// TIA Portal V19 export
FUNCTION_BLOCK "V20_BLOCK"   // FB40, LAD
{ S7_Optimized_Access := 'FALSE' }
// stored: SetENOAutomatically false
   VAR
      MB_LOAD { S7_SetPoint := 'True'} : Modbus_Comm_Load;
      MB_READ_ZSW { S7_SetPoint := 'True'} : Modbus_Master;
      MB_READ_HIW { S7_SetPoint := 'True'} : Modbus_Master;
      MB_WRITE_STW { S7_SetPoint := 'True'} : Modbus_Master;
      MB_WRITE_HSW { S7_SetPoint := 'True'} : Modbus_Master;
      DRIVE { S7_SetPoint := 'True'} : Array[1..11] of "VFD";
      DRIVE_ID { S7_SetPoint := 'True'} : Int := 1;
      STATUS : Int;
      MB_DB : P2P_MB_BASE;
      ZSW_DELAY { S7_SetPoint := 'True'} : TON_TIME;
      HIW_DELAY { S7_SetPoint := 'True'} : TON_TIME;
      STW_DELAY { S7_SetPoint := 'True'} : TON_TIME;
      HSW_DELAY { S7_SetPoint := 'True'} : TON_TIME;
      MB_READ_DI { S7_SetPoint := 'True'} : Modbus_Master;
      Modbus_Master_Instance { S7_SetPoint := 'True'} : Modbus_Master;
   END_VAR
   // DRIVE[1].ADDR := 1;
   // DRIVE[2].ADDR := 2;
   // DRIVE[3].ADDR := 3;
   // DRIVE[4].ADDR := 4;
   // DRIVE[5].ADDR := 5;
   // DRIVE[6].ADDR := 6;
   VAR_TEMP   // added for the SCL form of the ladder/FBD networks
      _w1 : Bool;
   END_VAR
BEGIN

REGION Network 1
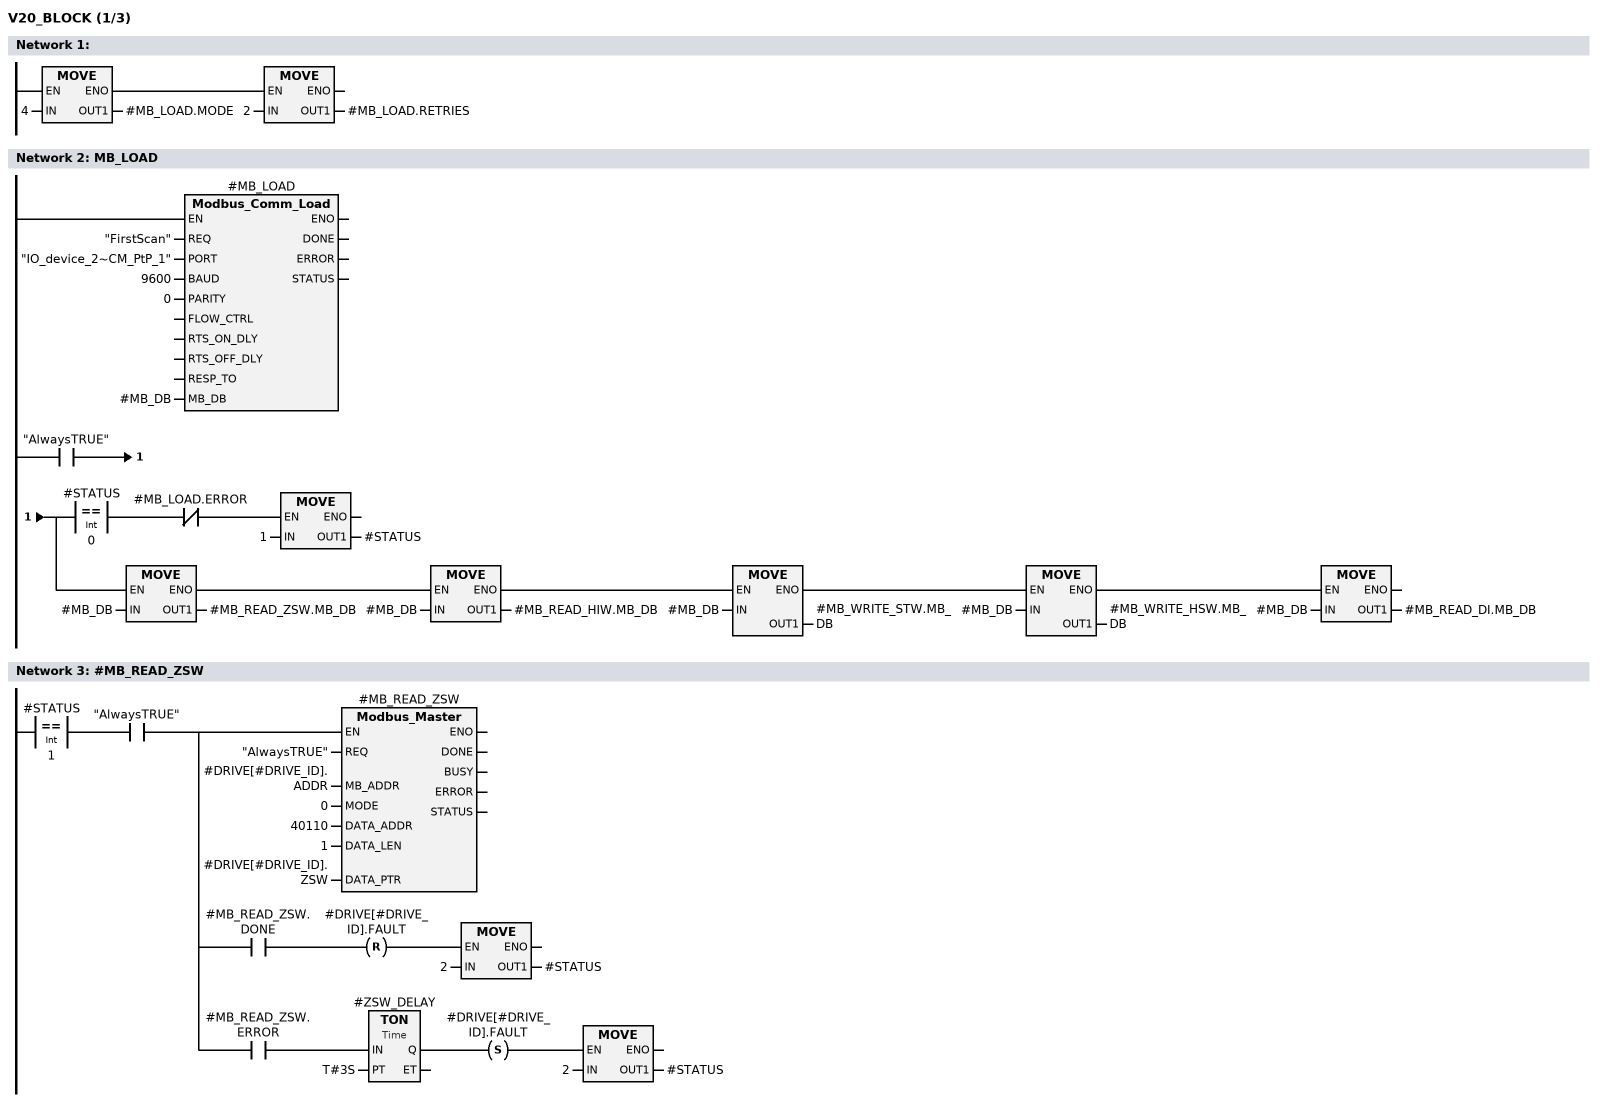
   RUNG wire#powerrail
      Move(in := 4, out1 => #MB_LOAD.MODE)
      Move(in := 2, out1 => #MB_LOAD.RETRIES)
   END_RUNG
   // the same network as SCL:
   #MB_LOAD.MODE := 4;
   #MB_LOAD.RETRIES := 2;
END_REGION

REGION Network 2: MB_LOAD
   RUNG wire#powerrail
      #MB_LOAD.Modbus_Comm_Load(REQ := "FirstScan", PORT := "IO_device_2~CM_PtP_1", BAUD := 9600, PARITY := 0, FLOW_CTRL :=, RTS_ON_DLY :=, RTS_OFF_DLY :=, RESP_TO :=, MB_DB := #MB_DB, DONE =>, ERROR =>, STATUS =>)
   END_RUNG
   RUNG wire#powerrail
      Contact( "AlwaysTRUE" )
      wire#w1
      { S7_Templates := "SrcType := Int" } EQ_Contact(in1 := #STATUS, in2 := 0)
      I_Contact( #MB_LOAD.ERROR )
      Move(in := 1, out1 => #STATUS)
   END_RUNG
   RUNG wire#w1
      Move(in := #MB_DB, out1 => #MB_READ_ZSW.MB_DB)
      Move(in := #MB_DB, out1 => #MB_READ_HIW.MB_DB)
      Move(in := #MB_DB, out1 => #MB_WRITE_STW.MB_DB)
      Move(in := #MB_DB, out1 => #MB_WRITE_HSW.MB_DB)
      Move(in := #MB_DB, out1 => #MB_READ_DI.MB_DB)
   END_RUNG
   // the same network as SCL:
   #MB_LOAD(REQ := "FirstScan", PORT := "IO_device_2~CM_PtP_1", BAUD := 9600, PARITY := 0, MB_DB := #MB_DB);   // Modbus_Comm_Load
   IF "AlwaysTRUE" AND (#STATUS = 0) AND NOT #MB_LOAD.ERROR THEN #STATUS := 1; END_IF;
   IF "AlwaysTRUE" THEN
       #MB_READ_ZSW.MB_DB := #MB_DB;
       #MB_READ_HIW.MB_DB := #MB_DB;
       #MB_WRITE_STW.MB_DB := #MB_DB;
       #MB_WRITE_HSW.MB_DB := #MB_DB;
       #MB_READ_DI.MB_DB := #MB_DB;
   END_IF;
END_REGION

REGION Network 3: #MB_READ_ZSW
   RUNG wire#powerrail
      { S7_Templates := "SrcType := Int" } EQ_Contact(in1 := #STATUS, in2 := 1)
      Contact( "AlwaysTRUE" )
      wire#w1
      #MB_READ_ZSW.Modbus_Master(REQ := "AlwaysTRUE", MB_ADDR := #DRIVE[#DRIVE_ID].ADDR, MODE := 0, DATA_ADDR := 40110, DATA_LEN := 1, DATA_PTR := #DRIVE[#DRIVE_ID].ZSW, DONE =>, BUSY =>, ERROR =>, STATUS =>)
   END_RUNG
   RUNG wire#w1
      Contact( #MB_READ_ZSW.DONE )
      R_Coil( #DRIVE[#DRIVE_ID].FAULT )
      Move(in := 2, out1 => #STATUS)
   END_RUNG
   RUNG wire#w1
      Contact( #MB_READ_ZSW.ERROR )
      { S7_Templates := "time_type := Time" } #ZSW_DELAY.TON(pt := T#3S, et =>)
      S_Coil( #DRIVE[#DRIVE_ID].FAULT )
      Move(in := 2, out1 => #STATUS)
   END_RUNG
   // the same network as SCL:
   #_w1 := (#STATUS = 1) AND "AlwaysTRUE";
   IF #_w1 THEN
       #MB_READ_ZSW(REQ := "AlwaysTRUE",   // Modbus_Master
                    MB_ADDR := #DRIVE[#DRIVE_ID].ADDR,
                    MODE := 0,
                    DATA_ADDR := 40110,
                    DATA_LEN := 1,
                    DATA_PTR := #DRIVE[#DRIVE_ID].ZSW);
   END_IF;
   IF #_w1 AND #MB_READ_ZSW.DONE THEN
       #DRIVE[#DRIVE_ID].FAULT := FALSE;
       #STATUS := 2;
   END_IF;
   #ZSW_DELAY(IN := #_w1 AND #MB_READ_ZSW.ERROR, PT := T#3S);   // TON
   IF #ZSW_DELAY.Q THEN
       #DRIVE[#DRIVE_ID].FAULT := TRUE;
       #STATUS := 2;
   END_IF;
END_REGION

REGION Network 4: #MB_READ_HIW
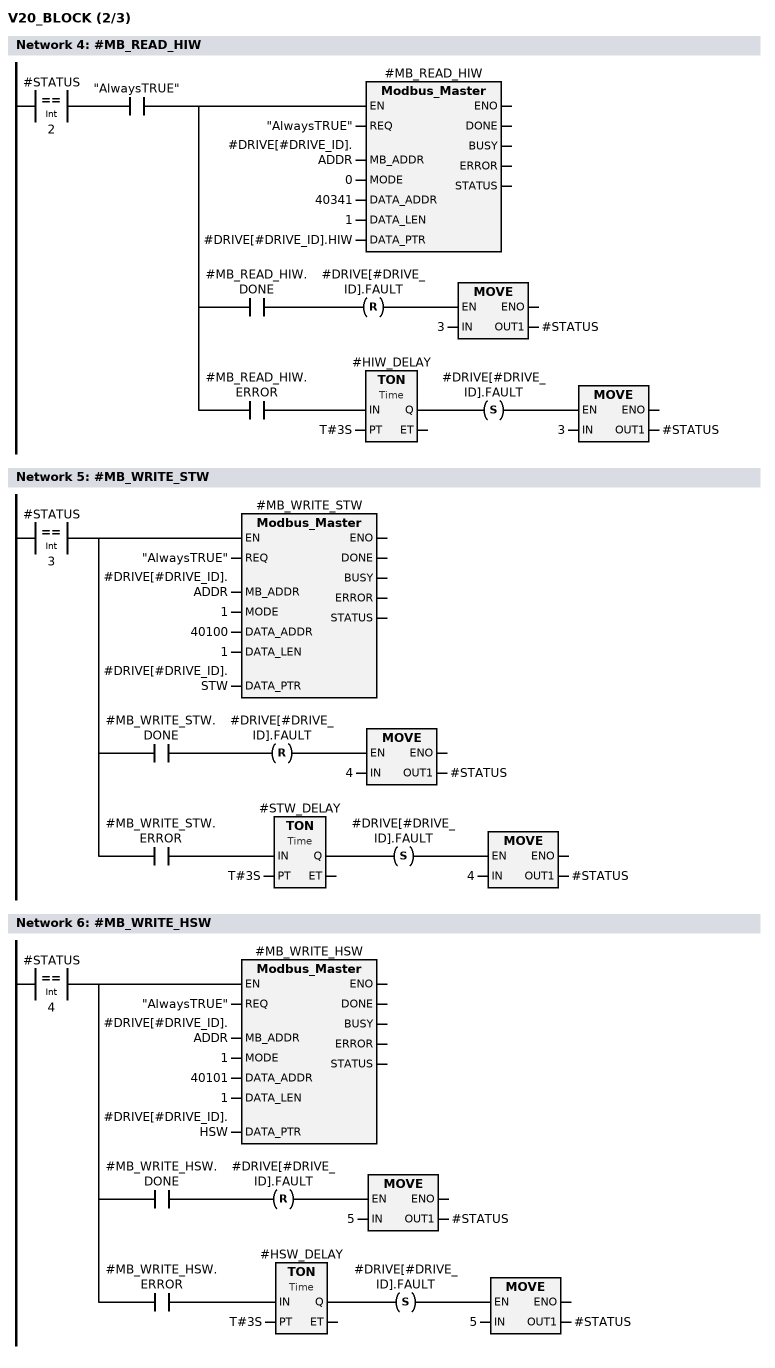
   RUNG wire#powerrail
      { S7_Templates := "SrcType := Int" } EQ_Contact(in1 := #STATUS, in2 := 2)
      Contact( "AlwaysTRUE" )
      wire#w1
      #MB_READ_HIW.Modbus_Master(REQ := "AlwaysTRUE", MB_ADDR := #DRIVE[#DRIVE_ID].ADDR, MODE := 0, DATA_ADDR := 40341, DATA_LEN := 1, DATA_PTR := #DRIVE[#DRIVE_ID].HIW, DONE =>, BUSY =>, ERROR =>, STATUS =>)
   END_RUNG
   RUNG wire#w1
      Contact( #MB_READ_HIW.DONE )
      R_Coil( #DRIVE[#DRIVE_ID].FAULT )
      Move(in := 3, out1 => #STATUS)
   END_RUNG
   RUNG wire#w1
      Contact( #MB_READ_HIW.ERROR )
      { S7_Templates := "time_type := Time" } #HIW_DELAY.TON(pt := T#3S, et =>)
      S_Coil( #DRIVE[#DRIVE_ID].FAULT )
      Move(in := 3, out1 => #STATUS)
   END_RUNG
   // the same network as SCL:
   #_w1 := (#STATUS = 2) AND "AlwaysTRUE";
   IF #_w1 THEN
       #MB_READ_HIW(REQ := "AlwaysTRUE",   // Modbus_Master
                    MB_ADDR := #DRIVE[#DRIVE_ID].ADDR,
                    MODE := 0,
                    DATA_ADDR := 40341,
                    DATA_LEN := 1,
                    DATA_PTR := #DRIVE[#DRIVE_ID].HIW);
   END_IF;
   IF #_w1 AND #MB_READ_HIW.DONE THEN
       #DRIVE[#DRIVE_ID].FAULT := FALSE;
       #STATUS := 3;
   END_IF;
   #HIW_DELAY(IN := #_w1 AND #MB_READ_HIW.ERROR, PT := T#3S);   // TON
   IF #HIW_DELAY.Q THEN
       #DRIVE[#DRIVE_ID].FAULT := TRUE;
       #STATUS := 3;
   END_IF;
END_REGION

REGION Network 5: #MB_WRITE_STW
   RUNG wire#powerrail
      { S7_Templates := "SrcType := Int" } EQ_Contact(in1 := #STATUS, in2 := 3)
      wire#w1
      #MB_WRITE_STW.Modbus_Master(REQ := "AlwaysTRUE", MB_ADDR := #DRIVE[#DRIVE_ID].ADDR, MODE := 1, DATA_ADDR := 40100, DATA_LEN := 1, DATA_PTR := #DRIVE[#DRIVE_ID].STW, DONE =>, BUSY =>, ERROR =>, STATUS =>)
   END_RUNG
   RUNG wire#w1
      Contact( #MB_WRITE_STW.DONE )
      R_Coil( #DRIVE[#DRIVE_ID].FAULT )
      Move(in := 4, out1 => #STATUS)
   END_RUNG
   RUNG wire#w1
      Contact( #MB_WRITE_STW.ERROR )
      { S7_Templates := "time_type := Time" } #STW_DELAY.TON(pt := T#3S, et =>)
      S_Coil( #DRIVE[#DRIVE_ID].FAULT )
      Move(in := 4, out1 => #STATUS)
   END_RUNG
   // the same network as SCL:
   #_w1 := #STATUS = 3;
   IF #_w1 THEN
       #MB_WRITE_STW(REQ := "AlwaysTRUE",   // Modbus_Master
                     MB_ADDR := #DRIVE[#DRIVE_ID].ADDR,
                     MODE := 1,
                     DATA_ADDR := 40100,
                     DATA_LEN := 1,
                     DATA_PTR := #DRIVE[#DRIVE_ID].STW);
   END_IF;
   IF #_w1 AND #MB_WRITE_STW.DONE THEN
       #DRIVE[#DRIVE_ID].FAULT := FALSE;
       #STATUS := 4;
   END_IF;
   #STW_DELAY(IN := #_w1 AND #MB_WRITE_STW.ERROR, PT := T#3S);   // TON
   IF #STW_DELAY.Q THEN
       #DRIVE[#DRIVE_ID].FAULT := TRUE;
       #STATUS := 4;
   END_IF;
END_REGION

REGION Network 6: #MB_WRITE_HSW
   RUNG wire#powerrail
      { S7_Templates := "SrcType := Int" } EQ_Contact(in1 := #STATUS, in2 := 4)
      wire#w1
      #MB_WRITE_HSW.Modbus_Master(REQ := "AlwaysTRUE", MB_ADDR := #DRIVE[#DRIVE_ID].ADDR, MODE := 1, DATA_ADDR := 40101, DATA_LEN := 1, DATA_PTR := #DRIVE[#DRIVE_ID].HSW, DONE =>, BUSY =>, ERROR =>, STATUS =>)
   END_RUNG
   RUNG wire#w1
      Contact( #MB_WRITE_HSW.DONE )
      R_Coil( #DRIVE[#DRIVE_ID].FAULT )
      Move(in := 5, out1 => #STATUS)
   END_RUNG
   RUNG wire#w1
      Contact( #MB_WRITE_HSW.ERROR )
      { S7_Templates := "time_type := Time" } #HSW_DELAY.TON(pt := T#3S, et =>)
      S_Coil( #DRIVE[#DRIVE_ID].FAULT )
      Move(in := 5, out1 => #STATUS)
   END_RUNG
   // the same network as SCL:
   #_w1 := #STATUS = 4;
   IF #_w1 THEN
       #MB_WRITE_HSW(REQ := "AlwaysTRUE",   // Modbus_Master
                     MB_ADDR := #DRIVE[#DRIVE_ID].ADDR,
                     MODE := 1,
                     DATA_ADDR := 40101,
                     DATA_LEN := 1,
                     DATA_PTR := #DRIVE[#DRIVE_ID].HSW);
   END_IF;
   IF #_w1 AND #MB_WRITE_HSW.DONE THEN
       #DRIVE[#DRIVE_ID].FAULT := FALSE;
       #STATUS := 5;
   END_IF;
   #HSW_DELAY(IN := #_w1 AND #MB_WRITE_HSW.ERROR, PT := T#3S);   // TON
   IF #HSW_DELAY.Q THEN
       #DRIVE[#DRIVE_ID].FAULT := TRUE;
       #STATUS := 5;
   END_IF;
END_REGION

REGION Network 7: #MB_READ_DI
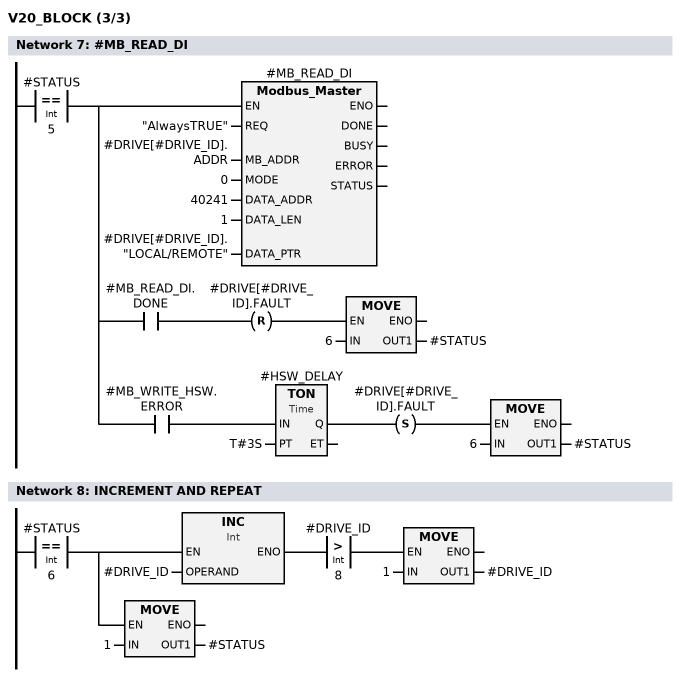
   RUNG wire#powerrail
      { S7_Templates := "SrcType := Int" } EQ_Contact(in1 := #STATUS, in2 := 5)
      wire#w1
      #MB_READ_DI.Modbus_Master(REQ := "AlwaysTRUE", MB_ADDR := #DRIVE[#DRIVE_ID].ADDR, MODE := 0, DATA_ADDR := 40241, DATA_LEN := 1, DATA_PTR := #DRIVE[#DRIVE_ID]."LOCAL/REMOTE", DONE =>, BUSY =>, ERROR =>, STATUS =>)
   END_RUNG
   RUNG wire#w1
      Contact( #MB_READ_DI.DONE )
      R_Coil( #DRIVE[#DRIVE_ID].FAULT )
      Move(in := 6, out1 => #STATUS)
   END_RUNG
   RUNG wire#w1
      Contact( #MB_WRITE_HSW.ERROR )
      { S7_Templates := "time_type := Time" } #HSW_DELAY.TON(pt := T#3S, et =>)
      S_Coil( #DRIVE[#DRIVE_ID].FAULT )
      Move(in := 6, out1 => #STATUS)
   END_RUNG
   // the same network as SCL:
   #_w1 := #STATUS = 5;
   IF #_w1 THEN
       #MB_READ_DI(REQ := "AlwaysTRUE",   // Modbus_Master
                   MB_ADDR := #DRIVE[#DRIVE_ID].ADDR,
                   MODE := 0,
                   DATA_ADDR := 40241,
                   DATA_LEN := 1,
                   DATA_PTR := #DRIVE[#DRIVE_ID]."LOCAL/REMOTE");
   END_IF;
   IF #_w1 AND #MB_READ_DI.DONE THEN
       #DRIVE[#DRIVE_ID].FAULT := FALSE;
       #STATUS := 6;
   END_IF;
   #HSW_DELAY(IN := #_w1 AND #MB_WRITE_HSW.ERROR, PT := T#3S);   // TON
   IF #HSW_DELAY.Q THEN
       #DRIVE[#DRIVE_ID].FAULT := TRUE;
       #STATUS := 6;
   END_IF;
END_REGION

REGION Network 8: INCREMENT AND REPEAT
   RUNG wire#powerrail
      { S7_Templates := "SrcType := Int" } EQ_Contact(in1 := #STATUS, in2 := 6)
      wire#w1
      { S7_Templates := "DestType := Int" } Inc( #DRIVE_ID )
      { S7_Templates := "SrcType := Int" } GT_Contact(in1 := #DRIVE_ID, in2 := 8)
      Move(in := 1, out1 => #DRIVE_ID)
   END_RUNG
   RUNG wire#w1
      Move(in := 1, out1 => #STATUS)
   END_RUNG
   // the same network as SCL:
   #_w1 := #STATUS = 6;
   IF #_w1 THEN #DRIVE_ID := #DRIVE_ID + 1; END_IF;
   IF #_w1 AND (#DRIVE_ID > 8) THEN #DRIVE_ID := 1; END_IF;
   IF #_w1 THEN #STATUS := 1; END_IF;
END_REGION
END_FUNCTION_BLOCK
